(* IEC 61131-3 sources: generating_plc_code_with_llms/Code#2/StableCode/third run, 10 files *)

(* ---- 10.st ---- *)
// 8.177951097488403s
// 1

// sigmoid function
function sigmoid(x) {
  var input = VAR_INPUT.X;
  END_VAR

  // code goes here...

  RETURN
}

(* ---- 11.st ---- *)
// 12.45738673210144s
// 2

//IEC 61131-3 sign function
function sign(x)
    VAR_INPUT
        y : INTEGER;
    END_VAR

    IF (x.GT. 0) THEN
        y = 1;
    ELSEIF (x.EQ. 0) THEN
        y = 0;
    ELSE
        y = -1;
    END IF

    RETURN y;
END function

(* ---- 13.st ---- *)
// 21.416545152664185s
// 2

// Function to select a random number from the list
FUNCTION SelectRandomNumber()

    // Initialize variables
    VAR
        nIndex : INTEGER;
        nRandNum : INTEGER;
    END_VAR

    // Generate random number between 0 and MAXNUMBERS
    nIndex = CONSTANT.MAXNUMBERS;
    WHILE (nIndex > 0) DO
        SET nIndex := nIndex - 1;
        nRandNum := CONSTANT.aNumbers[nIndex] MOD 256;
    END_WHILE

    // Check if the number 10 is found
    IF (nRandNum = 10) THEN
        ABORT;
    END_IF

    RETURN nRandNum;
END

(* ---- 15.st ---- *)
// 16.75307559967041s
// 1
public static void FC1002(OBJECT obj) {
    VAR_INPUT();
    VAR_IN_OUT();
    FUNCTION fc1002 :BOOL {
        E_A = TRUE;
        SENSOR = FALSE;
        ZEITW = TIME.CurrentTime;
        RETURN false;
    }
    END_FUNCTION
}

(* ---- 20.st ---- *)
// 21.822731971740723s
// 2
FUNCTION FUNCTION_BLOCK INTERLOCK()
    VAR_INPUT
        I1 : BOOL;
        I2 : BOOL;
        TL : TIME;
    END_VAR
    VAR_OUTPUT
        Q1 : BOOL;
        Q2 : BOOL;
    END_VAR
    VAR
        T1 : TOF;
        T2 : TOF;
    END_VAR

    IF (I1.AND. I2) THEN
        RETURN
    END_IF

    WAITFOR(TL)
    IF (I1.OR. I2) THEN
        Q1 := TRUE;
        Q2 := FALSE;
    ELSE
        Q1 := FALSE;
        Q2 := TRUE;
    END_IF
END FUNCTION

(* ---- 16.st ---- *)
// 22.658372163772583s
// 2
// Traffic Light Program in IEC 61131-3
// by J.K. Rowland

// Declare variables
VAR
    North_green : BOOL;
    North_yellow : BOOL;
    North_red : BOOL;
    East_green : BOOL;
    East_yellow : BOOL;
    East_red : BOOL;
    T1 : TON;
END_VAR

// Set up timer 1
T1.Init(10000);

// Traffic Light Control Structure
WHILE (T1.Read() > 0) DO
    IF North_green = TRUE THEN
        North_yellow = FALSE;
        North_red = FALSE;
    END IF;
    IF North_yellow = TRUE THEN
        North_red = FALSE;
    END IF;
    IF North_red = TRUE THEN
        East_green = FALSE;
        East_yellow = FALSE;
        East_red = FALSE;
    END IF;
    IF East_green = TRUE THEN
        East_yellow = FALSE;
        East_red = FALSE;
    END IF;
    IF East_yellow = TRUE THEN
        East_red = FALSE;
    END IF;
END WHILE;

(* ---- 17.st ---- *)
// 26.766207933425903s
// 2
// Declare Variables
INT aiOutside, aiHumidity;
STRING sShowText;

// Initialize Variables
aiOutside = 0;
aiHumidity = 0;
sShowText = "";

// Check Temperature and Display Text
IF (aiHumidity < 40 || (aiHumidity > 75 && aiOutside > 18) || aiOutside > 25) THEN
    sShowText := "Temp. OK";
ELSE IF (aiHumidity >= 40 && aiHumidity <= 75 && aiOutside > 18 && aiOutside < 25) THEN
    sShowText := "Opt";
ELSE
    sShowText := "Hot";
END_IF

// Display Result
Display.Message(sShowText);

(* ---- 4.st ---- *)
// 29.920950174331665s
// 2
// IEC 61131-3 Structured Text Program of a Fill Level Check
// fill level in a container should be monitored in three ranges: low, ok and high
// use one output each for low,ok and high
// the fill level is read in via an analog value (0 - 32767) and should be converted internally to 0-100%
IF aiLevel <= 32767 THEN
    PercentLevel = 100;
ELSE
    PercentLevel = (aiLevel * 100) / 32767;
END_IF
// check if the content falls below 1%
DO_IF(PercentLevel < 1)
    PlaySound("WarningHorn");
END_DO_IF
// solve this application by using CASE instruction
CASE PercentLevel
    WHEN 0 THEN
        doLow = TRUE;
    WHEN 25 THEN
        doOk = TRUE;
    WHEN 50 THEN
        doHigh = TRUE;
    WHEN 75 THEN
        doAlarm = TRUE;
    END_CASE

(* ---- 6.st ---- *)
// 66.72478818893433s
// 1
Give me an IEC 61131-3 structured text program of a crane lift. Two conveyor belts (doConvTop, doConvBottom) transport crate<s> to a lift. When the light barrier (diConvTop or diConvBottom) is activated, the corresponding conveyor belt stops and the lift is requested. If the lift has not yet been requested, it is moved to the corresponding position (doLiftTop, doLiftBottom). If the lift is in the requested position (diLiftTop, diLiftBottom), the lift conveyor belt (doConvLift) is switched on until the crate is completely at the lift (diBoxLift). The lift then moves to the unloading position (doLiftUnload). Once it has reached the position (diLiftUnload), the crate is the box is conveyeD onto the unloading conveyor. When the box has left the lift, it is free for the next request.
Following rules should be followed:
- variables should be declared between VAR and END_VAR
- when using control structures do not forget END_<controll structure>
- switch cases should be avoided unless instructed in the task
- use the right quotation marks for the string type
- implementing a function should be avoided
- only when implementing a function: the variables should be declared inside the function; the return value should be stored in a variable named after the function; RETURN should be used correctly, to return to the main method and not to return a value
Only following variables should be used:import java.util.*;

public class CraneLift {
    public static void main(String[] args) {
        VAR
            CONSTANT
                WAIT : UINT:= 0;
                TOP_POSITION : UINT:= 1;
                BOTTOM_POSITION : UINT:= 2;
                GETBOX : UINT:= 3;
                UNLOAD_POSITION : UINT:= 4;
                UNLOAD_BOX : UINT:= 5;
            END_VAR

            VAR
                (*-- digital outputs*)
                doConvTop: BOOL;
                doConvBottom: BOOL;
                doConvLift: BOOL;
                doLiftTop: BOOL;
                doLiftBottom: BOOL;
                doLiftUnload: BOOL;
                (*-- digital inputs*)
                diConvTop: BOOL;
                diConvBottom: BOOL;
                diLiftTop: BOOL;
                diLiftBottom: BOOL;
                diLiftUnload: BOOL;

(* ---- 8.st ---- *)
// 45.69720149040222s
// 1
procedure lambertW(varInput, var)
  VAR
    X : REAL;
  END_VAR

  VAR
    w : REAL;
    i : INT;
    we : REAL;
    w1e : REAL;
    ewx : REAL;
    last : DWORD;
  END_VAR

  begin

    for (i := 0 to 254) do
      begin
        X := varInput.real(i);
        w := lambertWValue(X);
        we := lambertWeValue(w, X);
        w1e := lambertWValue(we, X);
        ewx := lambertEwValue(w1e, X);
        last := i;
      end

    writeln("last = ", last);

  end procedure lambertW;

procedure lambertWValue(x, var)
  VAR
    w : REAL;
    x : REAL;
  END_VAR

  begin
    w := (2 * pi) * exp(-x**2 / 2);
  end procedure lambertWValue;

procedure lambertWeValue(w, var)
  VAR
    we : REAL;
    w : REAL;
    var : REAL;
  END_VAR

  begin
    we := sqrt((var**2 + (w*var)) / (var**2 + 1));
  end procedure lambertWeValue;

procedure lambertW1eValue(x, var)
  VAR
    w1e : REAL;
    x : REAL;
    var : REAL;
  END_VAR

  begin
    w1e := sqrt((var**2 + (w*var)) / (var**2 + 1));
  end procedure lambertW1eValue;

procedure lambertEwValue(w1e, var)
  VAR
    ewx : REAL;
    w1e : REAL;
    var : REAL;
  END_VAR

  begin
    ewx := sqrt((var**2 + (w*var)) / (var**2 + 1));
  end procedure lambertEwValue;
